(* IEC 61131-3 sources: llm-plc-st-eval/data/processed_v2_primera/claude-sonnet-4-6/I2/zero_shot, 3 files *)

(* ---- ejec_1.st ---- *)
FUNCTION_BLOCK FB_Llenado
VAR_INPUT
    nivelAlto  : BOOL; (* Sensor de nivel alto *)
    nivelBajo  : BOOL; (* Sensor de nivel bajo *)
    btnInicio  : BOOL; (* Botón de inicio (flanco o nivel) *)
    btnParo    : BOOL; (* Botón de paro (detiene todo) *)
END_VAR

VAR_OUTPUT
    vLlenado    : BOOL; (* Válvula de llenado *)
    motorMezcla : BOOL; (* Motor de mezcla *)
    vDescarga   : BOOL; (* Válvula de descarga *)
END_VAR

VAR
    (* Etapas del proceso *)
    eReposo    : BOOL := TRUE;  (* Etapa 0: reposo *)
    eLlenado   : BOOL := FALSE; (* Etapa 1: llenando *)
    eMezcla    : BOOL := FALSE; (* Etapa 2: mezclando *)
    eDescarga  : BOOL := FALSE; (* Etapa 3: descargando *)

    (* Temporizador para la mezcla *)
    tMezcla    : TON;
END_VAR

(* ─────────────────────────────────────────────
   PARO DE EMERGENCIA: tiene prioridad absoluta
   ───────────────────────────────────────────── *)
IF btnParo THEN
    (* Desactivar todas las salidas *)
    vLlenado    := FALSE;
    motorMezcla := FALSE;
    vDescarga   := FALSE;

    (* Resetear temporizador *)
    tMezcla(IN := FALSE, PT := T#60S);

    (* Volver a reposo *)
    eReposo  := TRUE;
    eLlenado := FALSE;
    eMezcla  := FALSE;
    eDescarga := FALSE;

ELSE
    (* ─────────────────────────────────────────
       ETAPA 0 – REPOSO
       ───────────────────────────────────────── *)
    IF eReposo THEN
        (* Todas las salidas apagadas *)
        vLlenado    := FALSE;
        motorMezcla := FALSE;
        vDescarga   := FALSE;

        (* Transición: btnInicio arranca el proceso *)
        IF btnInicio THEN
            eReposo  := FALSE;
            eLlenado := TRUE;
        END_IF;

    (* ─────────────────────────────────────────
       ETAPA 1 – LLENADO
       ───────────────────────────────────────── *)
    ELSIF eLlenado THEN
        vLlenado    := TRUE;  (* Abrir válvula de llenado *)
        motorMezcla := FALSE;
        vDescarga   := FALSE;

        (* Transición: nivel alto alcanzado *)
        IF nivelAlto THEN
            vLlenado := FALSE; (* Cerrar válvula antes de mezclar *)
            eLlenado := FALSE;
            eMezcla  := TRUE;
            tMezcla(IN := FALSE, PT := T#60S); (* Asegurar reset previo *)
        END_IF;

    (* ─────────────────────────────────────────
       ETAPA 2 – MEZCLA (60 s)
       ───────────────────────────────────────── *)
    ELSIF eMezcla THEN
        vLlenado    := FALSE;
        motorMezcla := TRUE;  (* Activar motor de mezcla *)
        vDescarga   := FALSE;

        (* Llamada al temporizador TON *)
        tMezcla(IN := TRUE, PT := T#60S);

        (* Transición: tiempo de mezcla cumplido *)
        IF tMezcla.Q THEN
            motorMezcla := FALSE;
            tMezcla(IN := FALSE, PT := T#60S); (* Resetear temporizador *)
            eMezcla   := FALSE;
            eDescarga := TRUE;
        END_IF;

    (* ─────────────────────────────────────────
       ETAPA 3 – DESCARGA
       ───────────────────────────────────────── *)
    ELSIF eDescarga THEN
        vLlenado    := FALSE;
        motorMezcla := FALSE;
        vDescarga   := TRUE;  (* Abrir válvula de descarga *)

        (* Transición: nivel bajo alcanzado (tanque vacío) *)
        IF nivelBajo THEN
            vDescarga := FALSE; (* Cerrar válvula *)
            eDescarga := FALSE;
            eReposo   := TRUE;  (* Volver a reposo *)
        END_IF;

    END_IF;

END_IF;

(* ---- ejec_2.st ---- *)
FUNCTION_BLOCK FB_Llenado
VAR_INPUT
    nivelAlto  : BOOL; (* Sensor de nivel alto *)
    nivelBajo  : BOOL; (* Sensor de nivel bajo *)
    btnInicio  : BOOL; (* Botón de inicio del proceso *)
    btnParo    : BOOL; (* Botón de paro de emergencia *)
END_VAR

VAR_OUTPUT
    vLlenado    : BOOL; (* Válvula de llenado *)
    motorMezcla : BOOL; (* Motor de mezcla *)
    vDescarga   : BOOL; (* Válvula de descarga *)
END_VAR

VAR
    (* Etapas del proceso *)
    etapa : INT := 0;
    (*
        0 = Reposo
        1 = Llenado
        2 = Mezcla
        3 = Descarga
    *)

    (* Temporizador para la etapa de mezcla *)
    tmrMezcla : TON;
END_VAR

(* ─────────────────────────────────────────────
   Lógica principal del proceso por etapas
   ───────────────────────────────────────────── *)

(* Paro de emergencia: cualquier etapa → reposo *)
IF btnParo THEN
    etapa       := 0;
    vLlenado    := FALSE;
    motorMezcla := FALSE;
    vDescarga   := FALSE;
    tmrMezcla(IN := FALSE); (* Reinicia el temporizador *)

ELSE

    CASE etapa OF

        (* ── Etapa 0: Reposo ── *)
        0:
            vLlenado    := FALSE;
            motorMezcla := FALSE;
            vDescarga   := FALSE;
            tmrMezcla(IN := FALSE); (* Mantiene temporizador reseteado *)

            IF btnInicio THEN
                etapa := 1; (* Ir a llenado *)
            END_IF;

        (* ── Etapa 1: Llenado ── *)
        1:
            vLlenado    := TRUE;
            motorMezcla := FALSE;
            vDescarga   := FALSE;

            IF nivelAlto THEN
                vLlenado := FALSE;
                etapa    := 2; (* Ir a mezcla *)
            END_IF;

        (* ── Etapa 2: Mezcla (60 segundos) ── *)
        2:
            vLlenado    := FALSE;
            motorMezcla := TRUE;
            vDescarga   := FALSE;

            (* Activa el temporizador mientras se está en esta etapa *)
            tmrMezcla(IN := TRUE, PT := T#60S);

            IF tmrMezcla.Q THEN
                motorMezcla := FALSE;
                tmrMezcla(IN := FALSE); (* Resetea para próximo ciclo *)
                etapa := 3;             (* Ir a descarga *)
            END_IF;

        (* ── Etapa 3: Descarga ── *)
        3:
            vLlenado    := FALSE;
            motorMezcla := FALSE;
            vDescarga   := TRUE;

            IF nivelBajo THEN
                vDescarga := FALSE;
                etapa     := 0; (* Volver a reposo *)
            END_IF;

        (* ── Estado no definido: forzar reposo ── *)
        ELSE
            etapa       := 0;
            vLlenado    := FALSE;
            motorMezcla := FALSE;
            vDescarga   := FALSE;

    END_CASE;

END_IF;

END_FUNCTION_BLOCK

(* ---- ejec_3.st ---- *)
FUNCTION_BLOCK FB_Llenado
VAR_INPUT
    nivelAlto  : BOOL; (* Sensor de nivel alto *)
    nivelBajo  : BOOL; (* Sensor de nivel bajo *)
    btnInicio  : BOOL; (* Botón de inicio (normalmente abierto) *)
    btnParo    : BOOL; (* Botón de paro  (normalmente abierto) *)
END_VAR

VAR_OUTPUT
    vLlenado    : BOOL; (* Válvula de llenado  *)
    motorMezcla : BOOL; (* Motor de mezcla     *)
    vDescarga   : BOOL; (* Válvula de descarga *)
END_VAR

VAR
    (* Etapas del proceso *)
    etapa : INT := 0;
    (*
        0 = Reposo
        1 = Llenado
        2 = Mezcla
        3 = Descarga
    *)

    (* Temporizador para la etapa de mezcla *)
    tmrMezcla : TON;
END_VAR

(* ─────────────────────────────────────────────
   Lógica de paro: tiene prioridad sobre todo
   ───────────────────────────────────────────── *)
IF btnParo THEN
    etapa       := 0;
    vLlenado    := FALSE;
    motorMezcla := FALSE;
    vDescarga   := FALSE;
    tmrMezcla(IN := FALSE); (* Reinicia el temporizador *)
    RETURN;                  (* Sale del bloque de función *)
END_IF;

(* ─────────────────────────────────────────────
   Máquina de estados por etapas
   ───────────────────────────────────────────── *)
CASE etapa OF

    (* ── ETAPA 0: Reposo ── *)
    0:
        vLlenado    := FALSE;
        motorMezcla := FALSE;
        vDescarga   := FALSE;
        tmrMezcla(IN := FALSE); (* Mantiene temporizador reseteado *)

        IF btnInicio THEN
            etapa := 1; (* Avanza a llenado *)
        END_IF;

    (* ── ETAPA 1: Llenado ── *)
    1:
        vLlenado    := TRUE;
        motorMezcla := FALSE;
        vDescarga   := FALSE;

        IF nivelAlto THEN
            vLlenado := FALSE;
            etapa    := 2; (* Avanza a mezcla *)
        END_IF;

    (* ── ETAPA 2: Mezcla (60 s) ── *)
    2:
        vLlenado    := FALSE;
        motorMezcla := TRUE;
        vDescarga   := FALSE;

        (* Activa el temporizador mientras se está en esta etapa *)
        tmrMezcla(IN := TRUE, PT := T#60S);

        IF tmrMezcla.Q THEN
            motorMezcla := FALSE;
            tmrMezcla(IN := FALSE); (* Reinicia para próximo ciclo *)
            etapa := 3;             (* Avanza a descarga *)
        END_IF;

    (* ── ETAPA 3: Descarga ── *)
    3:
        vLlenado    := FALSE;
        motorMezcla := FALSE;
        vDescarga   := TRUE;

        IF nivelBajo THEN
            vDescarga := FALSE;
            etapa     := 0; (* Regresa a reposo *)
        END_IF;

    (* ── Estado no definido: seguridad ── *)
    ELSE
        etapa       := 0;
        vLlenado    := FALSE;
        motorMezcla := FALSE;
        vDescarga   := FALSE;

END_CASE;
